ABB RAPID module: SpacedName.mod

MODULE MOD_SpacedName

PERS wobjdata rdkWObj := [FALSE, TRUE, "", [[0,0,0],[1,0,0,0]],[[0,0,0],[1,0,0,0]]];
PERS tooldata rdkTool := [TRUE,[[0,0,0],[1,0,0,0]],[6.8,[0,0,15],[1,0,0,0],0,0,0.005]];
VAR speeddata rdkSpeed := [500,500,500,500];
VAR zonedata rdkZone := z1;
VAR extjoint rdkExtax := [9E9,9E9,9E9,9E9,9E9,9E9];

PROC main_RoboDK()
	SpacedName;
	EXIT;
ENDPROC

PROC SpacedName()
	!Program generated by RoboDK v5.9.4 for ABB IRB 1600-8/1.45 on 26/10/2026 01:01:07
	!Using nominal kinematics.
	var robtarget crt;
	crt := CRobT(\Tool:=rdkTool, \WObj:=rdkWObj);
	rdkExtax := crt.extax;
	ConfJ \On;
	ConfL \Off;
	!Spaced body
ENDPROC

ENDMODULE
